TYPE ST_HmiCoversStatus :
STRUCT
	bPresent	: BOOL;
	bOpened		: BOOL;
	bClosed		: BOOL;
	bError		: BOOL;
END_STRUCT
END_TYPE

(* stored: Version 1.1.0.1, ProductVersion 3.1.4024.15
   DUT ST_HmiCoversStatus: Id {a501da17-f529-49a4-8cee-f871c9cf74e1} *)
